Staubli VAL3: main.pgx

program main()
begin
  close(tCurrentTool)
  pPointRx.config.shoulder = lefty
  pPointRx.config.elbow = epositive
  pPointRx.config.wrist = wpositive
  pPointRx2.config.shoulder = lefty
  pPointRx2.config.elbow = epositive
  pPointRx2.config.wrist = wpositive
  mCurrentSpeed.tvel = 100.00
  mCurrentSpeed.blend = joint
  mCurrentSpeed.reach = 0.010
  mCurrentSpeed.leave = 0.010
  // Program SubPick start
  call MoveLine(1077.300,-56.172,837.243,-146.156,25.288,-102.118)
  Output[7]=true

  waitEndMove()
  // Program SubPick end

end
